Universal Robots URScript: FaiChun_9 Jan_1_arc_1.script

def Machining2():
  # Default parameters:
  global speed_ms = 0.05
  global speed_rads = 0.75
  global accel_mss = 3
  global accel_radss = 1.2
  global blend_radius_m = 0.0003

  # Add subprograms here
  # Start of main program
  # Program generated by RoboDK v5.6.8 for UR10e on 13/01/2025 16:29:17
  # Using nominal kinematics.
  blend_radius_m = 0.0003
  speed_ms = 0.05
  # set_reference(p[0.325000, -0.070000, 0.000000, 0.000000, 0.000000, 0.000000])
  set_tcp(p[0.000000, 0.000000, 0.252000, 0.000000, 0.000000, 0.000000])
  # Show Tool
  movej([0.739676, -0.896584, -2.557623, -1.258182, 1.570796, 2.310473],accel_radss,speed_rads,0,blend_radius_m)
  movel([0.739676, -1.045549, -2.705771, -0.961069, 1.570796, 2.310473],accel_mss,speed_ms,0,blend_radius_m)
  #SetTool1
  #M_RunCode6
  #SetRPM60000
  speed_ms = 0.05
  #M_RunCode3
  movel([0.739676, -1.073443, -2.722043, -0.916902, 1.570796, 2.310473],accel_mss,speed_ms,0,blend_radius_m)
  speed_ms = 0.003
  movel([0.739676, -1.080869, -2.726059, -0.905462, 1.570796, 2.310473],accel_mss,speed_ms,0,blend_radius_m)
  speed_ms = 0.007
  movel([0.521026, -1.435757, -2.529573, -0.747059, 1.570796, 2.091823],accel_mss,speed_ms,0,blend_radius_m)
  movel([0.234867, -1.438478, -2.527424, -0.746487, 1.570796, 1.805663],accel_mss,speed_ms,0,blend_radius_m)
  movel([0.339201, -1.087620, -2.723617, -0.901152, 1.570796, 1.909998],accel_mss,speed_ms,0,blend_radius_m)
  movel([0.739676, -1.080869, -2.726059, -0.905462, 1.570796, 2.310473],accel_mss,speed_ms,0,blend_radius_m)
  speed_ms = 0.003
  movel([0.739676, -1.073443, -2.722043, -0.916902, 1.570796, 2.310473],accel_mss,speed_ms,0,blend_radius_m)
  speed_ms = 0.05
  movel([0.739676, -1.045549, -2.705771, -0.961069, 1.570796, 2.310473],accel_mss,speed_ms,0,blend_radius_m)
  #M_RunCode9
  movel([0.722285, -1.051564, -2.703686, -0.957139, 1.570796, 2.293082],accel_mss,speed_ms,0,blend_radius_m)
  #M_RunCode3
  movel([0.722285, -1.079477, -2.719883, -0.913030, 1.570796, 2.293082],accel_mss,speed_ms,0,blend_radius_m)
  speed_ms = 0.003
  movel([0.722285, -1.086903, -2.723879, -0.901608, 1.570796, 2.293082],accel_mss,speed_ms,0,blend_radius_m)
  speed_ms = 0.007
  movel([0.717716, -1.094057, -2.721252, -0.897081, 1.570796, 2.288512],accel_mss,speed_ms,0,blend_radius_m)
  movel([0.716212, -1.105701, -2.716877, -0.889811, 1.570796, 2.287008],accel_mss,speed_ms,0,blend_radius_m)
  movel([0.711055, -1.104499, -2.717334, -0.890556, 1.570796, 2.281852],accel_mss,speed_ms,0,blend_radius_m)
  movel([0.713896, -1.109311, -2.715495, -0.887583, 1.570796, 2.284692],accel_mss,speed_ms,0,blend_radius_m)
  movel([0.708427, -1.117848, -2.712180, -0.882361, 1.570796, 2.279223],accel_mss,speed_ms,0,blend_radius_m)
  movel([0.707812, -1.118809, -2.711802, -0.881778, 1.570796, 2.278608],accel_mss,speed_ms,0,blend_radius_m)
  movel([0.707378, -1.119487, -2.711535, -0.881367, 1.570796, 2.278174],accel_mss,speed_ms,0,blend_radius_m)
  movel([0.699793, -1.117779, -2.712207, -0.882403, 1.570796, 2.270589],accel_mss,speed_ms,0,blend_radius_m)
  movel([0.704152, -1.110893, -2.714886, -0.886610, 1.570796, 2.274948],accel_mss,speed_ms,0,blend_radius_m)
  movel([0.701466, -1.110302, -2.715114, -0.886973, 1.570796, 2.272262],accel_mss,speed_ms,0,blend_radius_m)
  movel([0.694884, -1.120745, -2.711039, -0.880605, 1.570796, 2.265680],accel_mss,speed_ms,0,blend_radius_m)
  movel([0.705120, -1.123018, -2.710138, -0.879233, 1.570796, 2.275917],accel_mss,speed_ms,0,blend_radius_m)
  movel([0.604989, -1.283325, -2.632898, -0.796166, 1.570796, 2.175785],accel_mss,speed_ms,0,blend_radius_m)
  movel([0.530205, -1.410064, -2.549311, -0.753014, 1.570796, 2.101001],accel_mss,speed_ms,0,blend_radius_m)
  movel([0.521929, -1.408991, -2.550114, -0.753284, 1.570796, 2.092726],accel_mss,speed_ms,0,blend_radius_m)
  movel([0.518334, -1.415415, -2.545281, -0.751692, 1.570796, 2.089130],accel_mss,speed_ms,0,blend_radius_m)
  movel([0.520473, -1.415684, -2.545078, -0.751627, 1.570796, 2.091269],accel_mss,speed_ms,0,blend_radius_m)
  movel([0.522841, -1.411466, -2.548259, -0.752664, 1.570796, 2.093637],accel_mss,speed_ms,0,blend_radius_m)
  movel([0.528942, -1.412267, -2.547657, -0.752465, 1.570796, 2.099738],accel_mss,speed_ms,0,blend_radius_m)
  movel([0.528547, -1.412961, -2.547135, -0.752293, 1.570796, 2.099343],accel_mss,speed_ms,0,blend_radius_m)
  movel([0.528364, -1.413282, -2.546893, -0.752214, 1.570796, 2.099160],accel_mss,speed_ms,0,blend_radius_m)
  movel([0.521314, -1.417954, -2.543354, -0.751080, 1.570796, 2.092111],accel_mss,speed_ms,0,blend_radius_m)
  movec([0.521009, -1.418498, -2.542941, -0.750950, 1.570796, 2.091805],[0.520704, -1.419040, -2.542527, -0.750821, 1.570796, 2.091500],accel_mss,speed_ms,blend_radius_m)
  movec([0.520399, -1.419584, -2.542113, -0.750692, 1.570796, 2.091195],[0.520094, -1.420127, -2.541698, -0.750564, 1.570796, 2.090890],accel_mss,speed_ms,blend_radius_m)
  movel([0.524182, -1.420660, -2.541290, -0.750438, 1.570796, 2.094978],accel_mss,speed_ms,0,blend_radius_m)
  movel([0.520710, -1.426805, -2.536563, -0.749022, 1.570796, 2.091507],accel_mss,speed_ms,0,blend_radius_m)
  movel([0.516647, -1.426280, -2.536969, -0.749140, 1.570796, 2.087443],accel_mss,speed_ms,0,blend_radius_m)
  movel([0.514345, -1.430404, -2.533767, -0.748218, 1.570796, 2.085141],accel_mss,speed_ms,0,blend_radius_m)
  movel([0.508328, -1.429667, -2.534341, -0.748381, 1.570796, 2.079124],accel_mss,speed_ms,0,blend_radius_m)
  movel([0.510606, -1.425534, -2.537545, -0.749310, 1.570796, 2.081402],accel_mss,speed_ms,0,blend_radius_m)
  movel([0.506209, -1.429417, -2.534536, -0.748437, 1.570796, 2.077005],accel_mss,speed_ms,0,blend_radius_m)
  movel([0.501142, -1.428840, -2.534984, -0.748565, 1.570796, 2.071939],accel_mss,speed_ms,0,blend_radius_m)
  movel([0.500651, -1.428783, -2.535029, -0.748578, 1.570796, 2.071447],accel_mss,speed_ms,0,blend_radius_m)
  movel([0.500157, -1.428731, -2.535069, -0.748589, 1.570796, 2.070953],accel_mss,speed_ms,0,blend_radius_m)
  movel([0.503495, -1.422587, -2.539814, -0.749988, 1.570796, 2.074291],accel_mss,speed_ms,0,blend_radius_m)
  movel([0.507609, -1.423054, -2.539455, -0.749880, 1.570796, 2.078405],accel_mss,speed_ms,0,blend_radius_m)
  movel([0.508797, -1.420891, -2.541114, -0.750384, 1.570796, 2.079593],accel_mss,speed_ms,0,blend_radius_m)
  movel([0.502532, -1.420185, -2.541654, -0.750550, 1.570796, 2.073328],accel_mss,speed_ms,0,blend_radius_m)
  movel([0.498030, -1.428499, -2.535249, -0.748641, 1.570796, 2.068827],accel_mss,speed_ms,0,blend_radius_m)
  movel([0.497523, -1.428447, -2.535290, -0.748653, 1.570796, 2.068319],accel_mss,speed_ms,0,blend_radius_m)
  movel([0.497042, -1.428395, -2.535329, -0.748664, 1.570796, 2.067838],accel_mss,speed_ms,0,blend_radius_m)
  movel([0.383251, -1.423074, -2.539440, -0.749875, 1.570796, 1.954047],accel_mss,speed_ms,0,blend_radius_m)
  movel([0.263080, -1.430856, -2.533414, -0.748118, 1.570796, 1.833877],accel_mss,speed_ms,0,blend_radius_m)
  movel([0.265517, -1.422588, -2.539813, -0.749988, 1.570796, 1.836314],accel_mss,speed_ms,0,blend_radius_m)
  movel([0.258622, -1.423422, -2.539172, -0.749794, 1.570796, 1.829418],accel_mss,speed_ms,0,blend_radius_m)
  movel([0.257999, -1.425574, -2.537514, -0.749301, 1.570796, 1.828796],accel_mss,speed_ms,0,blend_radius_m)
  movel([0.262529, -1.425022, -2.537940, -0.749427, 1.570796, 1.833326],accel_mss,speed_ms,0,blend_radius_m)
  movel([0.260738, -1.431127, -2.533203, -0.748059, 1.570796, 1.831534],accel_mss,speed_ms,0,blend_radius_m)
  movel([0.259655, -1.431256, -2.533102, -0.748031, 1.570796, 1.830452],accel_mss,speed_ms,0,blend_radius_m)
  movel([0.255252, -1.427829, -2.535769, -0.748791, 1.570796, 1.826048],accel_mss,speed_ms,0,blend_radius_m)
  movel([0.252906, -1.428125, -2.535539, -0.748725, 1.570796, 1.823702],accel_mss,speed_ms,0,blend_radius_m)
  movel([0.251743, -1.432228, -2.532342, -0.747818, 1.570796, 1.822539],accel_mss,speed_ms,0,blend_radius_m)
  movel([0.245076, -1.433089, -2.531668, -0.747631, 1.570796, 1.815873],accel_mss,speed_ms,0,blend_radius_m)
  movel([0.246206, -1.428996, -2.534863, -0.748530, 1.570796, 1.817002],accel_mss,speed_ms,0,blend_radius_m)
  movel([0.243345, -1.423504, -2.539109, -0.749776, 1.570796, 1.814141],accel_mss,speed_ms,0,blend_radius_m)
  movel([0.247902, -1.422884, -2.539586, -0.749919, 1.570796, 1.818698],accel_mss,speed_ms,0,blend_radius_m)
  movel([0.248502, -1.420729, -2.541238, -0.750422, 1.570796, 1.819298],accel_mss,speed_ms,0,blend_radius_m)
  movel([0.243934, -1.421351, -2.540762, -0.750276, 1.570796, 1.814730],accel_mss,speed_ms,0,blend_radius_m)
  movel([0.245350, -1.416182, -2.544701, -0.751507, 1.570796, 1.816147],accel_mss,speed_ms,0,blend_radius_m)
  movel([0.252445, -1.414242, -2.546169, -0.751979, 1.570796, 1.823242],accel_mss,speed_ms,0,blend_radius_m)
  movel([0.251262, -1.418432, -2.542991, -0.750966, 1.570796, 1.822058],accel_mss,speed_ms,0,blend_radius_m)
  movel([0.253639, -1.418118, -2.543230, -0.751041, 1.570796, 1.824436],accel_mss,speed_ms,0,blend_radius_m)
  movel([0.255455, -1.411739, -2.548054, -0.752596, 1.570796, 1.826251],accel_mss,speed_ms,0,blend_radius_m)
  movel([0.246231, -1.412992, -2.547111, -0.752286, 1.570796, 1.817027],accel_mss,speed_ms,0,blend_radius_m)
  movel([0.282412, -1.287409, -2.630540, -0.794439, 1.570796, 1.853209],accel_mss,speed_ms,0,blend_radius_m)
  movel([0.331289, -1.130759, -2.707034, -0.874596, 1.570796, 1.902085],accel_mss,speed_ms,0,blend_radius_m)
  movel([0.331811, -1.129158, -2.707681, -0.875550, 1.570796, 1.902607],accel_mss,speed_ms,0,blend_radius_m)
  movel([0.344365, -1.126524, -2.708739, -0.877125, 1.570796, 1.915161],accel_mss,speed_ms,0,blend_radius_m)
  movel([0.347816, -1.116232, -2.712812, -0.883345, 1.570796, 1.918612],accel_mss,speed_ms,0,blend_radius_m)
  movel([0.344526, -1.116917, -2.712545, -0.882928, 1.570796, 1.915323],accel_mss,speed_ms,0,blend_radius_m)
  movel([0.342270, -1.123698, -2.709868, -0.878823, 1.570796, 1.913066],accel_mss,speed_ms,0,blend_radius_m)
  movel([0.332951, -1.125669, -2.709082, -0.877638, 1.570796, 1.903747],accel_mss,speed_ms,0,blend_radius_m)
  movel([0.333474, -1.124054, -2.709726, -0.878609, 1.570796, 1.904271],accel_mss,speed_ms,0,blend_radius_m)
  movel([0.342570, -1.114276, -2.713575, -0.884538, 1.570796, 1.913366],accel_mss,speed_ms,0,blend_radius_m)
  movel([0.343748, -1.110711, -2.714956, -0.886722, 1.570796, 1.914545],accel_mss,speed_ms,0,blend_radius_m)
  movel([0.340718, -1.101853, -2.718336, -0.892200, 1.570796, 1.911515],accel_mss,speed_ms,0,blend_radius_m)
  movel([0.347166, -1.100432, -2.718872, -0.893085, 1.570796, 1.917962],accel_mss,speed_ms,0,blend_radius_m)
  movel([0.349516, -1.093391, -2.721498, -0.897500, 1.570796, 1.920312],accel_mss,speed_ms,0,blend_radius_m)
  movel([0.359125, -1.091319, -2.722262, -0.898808, 1.570796, 1.929921],accel_mss,speed_ms,0,blend_radius_m)
  movel([0.356708, -1.098395, -2.719636, -0.894358, 1.570796, 1.927504],accel_mss,speed_ms,0,blend_radius_m)
  movec([0.357543, -1.098221, -2.719701, -0.894467, 1.570796, 1.928339],[0.358378, -1.098047, -2.719766, -0.894576, 1.570796, 1.929174],accel_mss,speed_ms,blend_radius_m)
  movec([0.359213, -1.097874, -2.719831, -0.894684, 1.570796, 1.930010],[0.360048, -1.097701, -2.719896, -0.894792, 1.570796, 1.930844],accel_mss,speed_ms,blend_radius_m)
  movel([0.362489, -1.090612, -2.722522, -0.899255, 1.570796, 1.933285],accel_mss,speed_ms,0,blend_radius_m)
  movel([0.372081, -1.088653, -2.723240, -0.900496, 1.570796, 1.942877],accel_mss,speed_ms,0,blend_radius_m)
  movel([0.368381, -1.099168, -2.719347, -0.893875, 1.570796, 1.939178],accel_mss,speed_ms,0,blend_radius_m)
  movel([0.361972, -1.100448, -2.718866, -0.893075, 1.570796, 1.932768],accel_mss,speed_ms,0,blend_radius_m)
  movel([0.360716, -1.104083, -2.717492, -0.890814, 1.570796, 1.931512],accel_mss,speed_ms,0,blend_radius_m)
  movel([0.370416, -1.102170, -2.718216, -0.892002, 1.570796, 1.941212],accel_mss,speed_ms,0,blend_radius_m)
  movel([0.375438, -1.087987, -2.723483, -0.900919, 1.570796, 1.946234],accel_mss,speed_ms,0,blend_radius_m)
  movel([0.546051, -1.068879, -2.730296, -0.913214, 1.570796, 2.116847],accel_mss,speed_ms,0,blend_radius_m)
  movel([0.701149, -1.082254, -2.725561, -0.904574, 1.570796, 2.271946],accel_mss,speed_ms,0,blend_radius_m)
  movel([0.692244, -1.096648, -2.720289, -0.895452, 1.570796, 2.263040],accel_mss,speed_ms,0,blend_radius_m)
  movel([0.700259, -1.098274, -2.719681, -0.894433, 1.570796, 2.271055],accel_mss,speed_ms,0,blend_radius_m)
  movel([0.702567, -1.094590, -2.721054, -0.896745, 1.570796, 2.273363],accel_mss,speed_ms,0,blend_radius_m)
  movel([0.697284, -1.093499, -2.721458, -0.897432, 1.570796, 2.268081],accel_mss,speed_ms,0,blend_radius_m)
  movel([0.703923, -1.082833, -2.725353, -0.904204, 1.570796, 2.274720],accel_mss,speed_ms,0,blend_radius_m)
  movel([0.704189, -1.082887, -2.725333, -0.904169, 1.570796, 2.274985],accel_mss,speed_ms,0,blend_radius_m)
  movel([0.705203, -1.083098, -2.725257, -0.904034, 1.570796, 2.275999],accel_mss,speed_ms,0,blend_radius_m)
  movel([0.711781, -1.084505, -2.724749, -0.903135, 1.570796, 2.282578],accel_mss,speed_ms,0,blend_radius_m)
  movel([0.707252, -1.091700, -2.722122, -0.898567, 1.570796, 2.278048],accel_mss,speed_ms,0,blend_radius_m)
  movel([0.709979, -1.092296, -2.721902, -0.898191, 1.570796, 2.280775],accel_mss,speed_ms,0,blend_radius_m)
  movel([0.722285, -1.086903, -2.723879, -0.901608, 1.570796, 2.293082],accel_mss,speed_ms,0,blend_radius_m)
  speed_ms = 0.003
  movel([0.722285, -1.079477, -2.719883, -0.913030, 1.570796, 2.293082],accel_mss,speed_ms,0,blend_radius_m)
  speed_ms = 0.05
  movel([0.722285, -1.051564, -2.703686, -0.957139, 1.570796, 2.293082],accel_mss,speed_ms,0,blend_radius_m)
  #M_RunCode9
  movel([0.397634, -1.094593, -2.687861, -0.929935, 1.570796, 1.968430],accel_mss,speed_ms,0,blend_radius_m)
  #M_RunCode3
  movel([0.397634, -1.122537, -2.703510, -0.886342, 1.570796, 1.968430],accel_mss,speed_ms,0,blend_radius_m)
  speed_ms = 0.003
  movel([0.397634, -1.129941, -2.707365, -0.875083, 1.570796, 1.968430],accel_mss,speed_ms,0,blend_radius_m)
  speed_ms = 0.007
  movec([0.397337, -1.130959, -2.706953, -0.874477, 1.570796, 1.968133],[0.396949, -1.131993, -2.706534, -0.873862, 1.570796, 1.967745],accel_mss,speed_ms,blend_radius_m)
  movec([0.396255, -1.133449, -2.705942, -0.872998, 1.570796, 1.967051],[0.395394, -1.134891, -2.705353, -0.872144, 1.570796, 1.966190],accel_mss,speed_ms,blend_radius_m)
  movec([0.394595, -1.136025, -2.704889, -0.871475, 1.570796, 1.965391],[0.393717, -1.137121, -2.704440, -0.870829, 1.570796, 1.964513],accel_mss,speed_ms,blend_radius_m)
  movec([0.392871, -1.138072, -2.704048, -0.870269, 1.570796, 1.963667],[0.391984, -1.138986, -2.703672, -0.869732, 1.570796, 1.962780],accel_mss,speed_ms,blend_radius_m)
  movec([0.390895, -1.140016, -2.703246, -0.869127, 1.570796, 1.961691],[0.389771, -1.140994, -2.702841, -0.868555, 1.570796, 1.960567],accel_mss,speed_ms,blend_radius_m)
  movec([0.388667, -1.141870, -2.702477, -0.868042, 1.570796, 1.959464],[0.387540, -1.142678, -2.702141, -0.867570, 1.570796, 1.958336],accel_mss,speed_ms,blend_radius_m)
  movec([0.386309, -1.143464, -2.701813, -0.867112, 1.570796, 1.957105],[0.385068, -1.144158, -2.701523, -0.866707, 1.570796, 1.955864],accel_mss,speed_ms,blend_radius_m)
  movel([0.384283, -1.144545, -2.701362, -0.866482, 1.570796, 1.955080],accel_mss,speed_ms,0,blend_radius_m)
  movec([0.382774, -1.145210, -2.701083, -0.866096, 1.570796, 1.953570],[0.381275, -1.145785, -2.700842, -0.865762, 1.570796, 1.952072],accel_mss,speed_ms,blend_radius_m)
  movec([0.379746, -1.146284, -2.700633, -0.865472, 1.570796, 1.950543],[0.378243, -1.146680, -2.700466, -0.865242, 1.570796, 1.949039],accel_mss,speed_ms,blend_radius_m)
  movel([0.377080, -1.146932, -2.700360, -0.865097, 1.570796, 1.947876],accel_mss,speed_ms,0,blend_radius_m)
  movec([0.375723, -1.147196, -2.700249, -0.864943, 1.570796, 1.946520],[0.374377, -1.147434, -2.700149, -0.864806, 1.570796, 1.945173],accel_mss,speed_ms,blend_radius_m)
  movec([0.372777, -1.147687, -2.700043, -0.864660, 1.570796, 1.943574],[0.371187, -1.147915, -2.699946, -0.864527, 1.570796, 1.941984],accel_mss,speed_ms,blend_radius_m)
  movec([0.368942, -1.148277, -2.699794, -0.864318, 1.570796, 1.939738],[0.366679, -1.148691, -2.699619, -0.864079, 1.570796, 1.937475],accel_mss,speed_ms,blend_radius_m)
  movec([0.365810, -1.148867, -2.699545, -0.863977, 1.570796, 1.936606],[0.364936, -1.149059, -2.699464, -0.863867, 1.570796, 1.935733],accel_mss,speed_ms,blend_radius_m)
  movel([0.364507, -1.149159, -2.699421, -0.863809, 1.570796, 1.935303],accel_mss,speed_ms,0,blend_radius_m)
  movec([0.363623, -1.149389, -2.699324, -0.863676, 1.570796, 1.934419],[0.362729, -1.149654, -2.699212, -0.863523, 1.570796, 1.933525],accel_mss,speed_ms,blend_radius_m)
  movec([0.361556, -1.150059, -2.699040, -0.863290, 1.570796, 1.932352],[0.360373, -1.150529, -2.698841, -0.863019, 1.570796, 1.931169],accel_mss,speed_ms,blend_radius_m)
  movel([0.359060, -1.151121, -2.698590, -0.862678, 1.570796, 1.929857],accel_mss,speed_ms,0,blend_radius_m)
  movel([0.357816, -1.151769, -2.698314, -0.862306, 1.570796, 1.928612],accel_mss,speed_ms,0,blend_radius_m)
  movec([0.356426, -1.152631, -2.697947, -0.861811, 1.570796, 1.927223],[0.355071, -1.153621, -2.697525, -0.861244, 1.570796, 1.925867],accel_mss,speed_ms,blend_radius_m)
  movec([0.354412, -1.154159, -2.697294, -0.860936, 1.570796, 1.925208],[0.353768, -1.154723, -2.697053, -0.860613, 1.570796, 1.924564],accel_mss,speed_ms,blend_radius_m)
  movel([0.353988, -1.155027, -2.696922, -0.860439, 1.570796, 1.924784],accel_mss,speed_ms,0,blend_radius_m)
  movel([0.354205, -1.155333, -2.696791, -0.860265, 1.570796, 1.925001],accel_mss,speed_ms,0,blend_radius_m)
  movel([0.354363, -1.155556, -2.696696, -0.860137, 1.570796, 1.925159],accel_mss,speed_ms,0,blend_radius_m)
  movec([0.355113, -1.156538, -2.696274, -0.859578, 1.570796, 1.925909],[0.355924, -1.157459, -2.695877, -0.859053, 1.570796, 1.926721],accel_mss,speed_ms,blend_radius_m)
  movec([0.356629, -1.158142, -2.695582, -0.858665, 1.570796, 1.927425],[0.357388, -1.158766, -2.695312, -0.858310, 1.570796, 1.928184],accel_mss,speed_ms,blend_radius_m)
  movec([0.358002, -1.159195, -2.695127, -0.858067, 1.570796, 1.928799],[0.358655, -1.159578, -2.694961, -0.857850, 1.570796, 1.929451],accel_mss,speed_ms,blend_radius_m)
  movec([0.359290, -1.159888, -2.694826, -0.857674, 1.570796, 1.930086],[0.359960, -1.160152, -2.694712, -0.857525, 1.570796, 1.930756],accel_mss,speed_ms,blend_radius_m)
  movec([0.360746, -1.160381, -2.694612, -0.857396, 1.570796, 1.931543],[0.361580, -1.160537, -2.694545, -0.857308, 1.570796, 1.932376],accel_mss,speed_ms,blend_radius_m)
  movel([0.362491, -1.160615, -2.694511, -0.857263, 1.570796, 1.933287],accel_mss,speed_ms,0,blend_radius_m)
  movec([0.363505, -1.160603, -2.694516, -0.857270, 1.570796, 1.934301],[0.364559, -1.160501, -2.694560, -0.857328, 1.570796, 1.935355],accel_mss,speed_ms,blend_radius_m)
  movec([0.365638, -1.160307, -2.694644, -0.857437, 1.570796, 1.936435],[0.366749, -1.160013, -2.694772, -0.857604, 1.570796, 1.937545],accel_mss,speed_ms,blend_radius_m)
  movec([0.368362, -1.159420, -2.695029, -0.857940, 1.570796, 1.939159],[0.369995, -1.158626, -2.695373, -0.858390, 1.570796, 1.940791],accel_mss,speed_ms,blend_radius_m)
  movec([0.371113, -1.157977, -2.695653, -0.858759, 1.570796, 1.941909],[0.372219, -1.157253, -2.695966, -0.859170, 1.570796, 1.943015],accel_mss,speed_ms,blend_radius_m)
  movel([0.360789, -1.167387, -2.691545, -0.853457, 1.570796, 1.931585],accel_mss,speed_ms,0,blend_radius_m)
  movel([0.344914, -1.145108, -2.701126, -0.866155, 1.570796, 1.915710],accel_mss,speed_ms,0,blend_radius_m)
  movel([0.346071, -1.144040, -2.701573, -0.866776, 1.570796, 1.916867],accel_mss,speed_ms,0,blend_radius_m)
  movec([0.347403, -1.142893, -2.702051, -0.867445, 1.570796, 1.918199],[0.348790, -1.141858, -2.702482, -0.868049, 1.570796, 1.919586],accel_mss,speed_ms,blend_radius_m)
  movec([0.349938, -1.141112, -2.702792, -0.868485, 1.570796, 1.920734],[0.351098, -1.140448, -2.703067, -0.868874, 1.570796, 1.921894],accel_mss,speed_ms,blend_radius_m)
  movec([0.351876, -1.140050, -2.703232, -0.869107, 1.570796, 1.922673],[0.352654, -1.139687, -2.703382, -0.869320, 1.570796, 1.923450],accel_mss,speed_ms,blend_radius_m)
  movec([0.354924, -1.138754, -2.703767, -0.869868, 1.570796, 1.925721],[0.357169, -1.137991, -2.704082, -0.870316, 1.570796, 1.927965],accel_mss,speed_ms,blend_radius_m)
  movec([0.358472, -1.137621, -2.704234, -0.870534, 1.570796, 1.929269],[0.359759, -1.137311, -2.704362, -0.870717, 1.570796, 1.930556],accel_mss,speed_ms,blend_radius_m)
  movec([0.360451, -1.137162, -2.704423, -0.870805, 1.570796, 1.931247],[0.361141, -1.137017, -2.704482, -0.870890, 1.570796, 1.931938],accel_mss,speed_ms,blend_radius_m)
  movec([0.362865, -1.136681, -2.704620, -0.871088, 1.570796, 1.933661],[0.364580, -1.136371, -2.704747, -0.871271, 1.570796, 1.935376],accel_mss,speed_ms,blend_radius_m)
  movec([0.366768, -1.136001, -2.704899, -0.871489, 1.570796, 1.937564],[0.368948, -1.135654, -2.705041, -0.871694, 1.570796, 1.939744],accel_mss,speed_ms,blend_radius_m)
  movec([0.371841, -1.135226, -2.705217, -0.871947, 1.570796, 1.942637],[0.374749, -1.134761, -2.705407, -0.872222, 1.570796, 1.945545],accel_mss,speed_ms,blend_radius_m)
  movec([0.375820, -1.134576, -2.705482, -0.872331, 1.570796, 1.946616],[0.376896, -1.134377, -2.705563, -0.872449, 1.570796, 1.947692],accel_mss,speed_ms,blend_radius_m)
  movel([0.377425, -1.134273, -2.705606, -0.872510, 1.570796, 1.948222],accel_mss,speed_ms,0,blend_radius_m)
  movec([0.379248, -1.133855, -2.705776, -0.872758, 1.570796, 1.950044],[0.381104, -1.133317, -2.705996, -0.873076, 1.570796, 1.951900],accel_mss,speed_ms,blend_radius_m)
  movec([0.382534, -1.132825, -2.706196, -0.873368, 1.570796, 1.953331],[0.383978, -1.132256, -2.706427, -0.873706, 1.570796, 1.954775],accel_mss,speed_ms,blend_radius_m)
  movec([0.385185, -1.131706, -2.706650, -0.874032, 1.570796, 1.955982],[0.386396, -1.131064, -2.706911, -0.874414, 1.570796, 1.957192],accel_mss,speed_ms,blend_radius_m)
  movec([0.387452, -1.130417, -2.707172, -0.874799, 1.570796, 1.958248],[0.388493, -1.129686, -2.707468, -0.875235, 1.570796, 1.959289],accel_mss,speed_ms,blend_radius_m)
  movec([0.389177, -1.129152, -2.707683, -0.875554, 1.570796, 1.959973],[0.389847, -1.128585, -2.707912, -0.875892, 1.570796, 1.960643],accel_mss,speed_ms,blend_radius_m)
  movec([0.390510, -1.127977, -2.708156, -0.876256, 1.570796, 1.961306],[0.391154, -1.127344, -2.708410, -0.876634, 1.570796, 1.961951],accel_mss,speed_ms,blend_radius_m)
  movel([0.392177, -1.126228, -2.708858, -0.877303, 1.570796, 1.962973],accel_mss,speed_ms,0,blend_radius_m)
  movel([0.393116, -1.125005, -2.709347, -0.878037, 1.570796, 1.963912],accel_mss,speed_ms,0,blend_radius_m)
  movel([0.393830, -1.123845, -2.709809, -0.878734, 1.570796, 1.964626],accel_mss,speed_ms,0,blend_radius_m)
  movel([0.394302, -1.122851, -2.710205, -0.879333, 1.570796, 1.965098],accel_mss,speed_ms,0,blend_radius_m)
  movel([0.394449, -1.122460, -2.710360, -0.879569, 1.570796, 1.965245],accel_mss,speed_ms,0,blend_radius_m)
  movec([0.394689, -1.121685, -2.710667, -0.880037, 1.570796, 1.965485],[0.394858, -1.120928, -2.710966, -0.880494, 1.570796, 1.965654],accel_mss,speed_ms,blend_radius_m)
  movec([0.394959, -1.119764, -2.711426, -0.881199, 1.570796, 1.965755],[0.394824, -1.118725, -2.711835, -0.881829, 1.570796, 1.965621],accel_mss,speed_ms,blend_radius_m)
  movel([0.394458, -1.117809, -2.712195, -0.882385, 1.570796, 1.965254],accel_mss,speed_ms,0,blend_radius_m)
  movec([0.394177, -1.117385, -2.712361, -0.882643, 1.570796, 1.964973],[0.393846, -1.117007, -2.712509, -0.882872, 1.570796, 1.964643],accel_mss,speed_ms,blend_radius_m)
  movel([0.393215, -1.116570, -2.712680, -0.883139, 1.570796, 1.964012],accel_mss,speed_ms,0,blend_radius_m)
  movel([0.392747, -1.116425, -2.712737, -0.883227, 1.570796, 1.963544],accel_mss,speed_ms,0,blend_radius_m)
  movel([0.392465, -1.116395, -2.712749, -0.883245, 1.570796, 1.963261],accel_mss,speed_ms,0,blend_radius_m)
  movel([0.391761, -1.116466, -2.712721, -0.883202, 1.570796, 1.962558],accel_mss,speed_ms,0,blend_radius_m)
  movel([0.391189, -1.116670, -2.712641, -0.883078, 1.570796, 1.961986],accel_mss,speed_ms,0,blend_radius_m)
  movel([0.390941, -1.116802, -2.712590, -0.882998, 1.570796, 1.961738],accel_mss,speed_ms,0,blend_radius_m)
  movel([0.390599, -1.117028, -2.712501, -0.882860, 1.570796, 1.961395],accel_mss,speed_ms,0,blend_radius_m)
  movel([0.390249, -1.117314, -2.712389, -0.882686, 1.570796, 1.961045],accel_mss,speed_ms,0,blend_radius_m)
  movel([0.390069, -1.117494, -2.712318, -0.882576, 1.570796, 1.960865],accel_mss,speed_ms,0,blend_radius_m)
  movel([0.389660, -1.118019, -2.712112, -0.882257, 1.570796, 1.960456],accel_mss,speed_ms,0,blend_radius_m)
  movel([0.389214, -1.118739, -2.711829, -0.881820, 1.570796, 1.960010],accel_mss,speed_ms,0,blend_radius_m)
  movel([0.389063, -1.119009, -2.711723, -0.881657, 1.570796, 1.959860],accel_mss,speed_ms,0,blend_radius_m)
  movel([0.388430, -1.120085, -2.711299, -0.881004, 1.570796, 1.959226],accel_mss,speed_ms,0,blend_radius_m)
  movel([0.388001, -1.120712, -2.711052, -0.880625, 1.570796, 1.958798],accel_mss,speed_ms,0,blend_radius_m)
  movel([0.387698, -1.121101, -2.710898, -0.880390, 1.570796, 1.958494],accel_mss,speed_ms,0,blend_radius_m)
  movel([0.386944, -1.121913, -2.710577, -0.879899, 1.570796, 1.957740],accel_mss,speed_ms,0,blend_radius_m)
  movel([0.385868, -1.122888, -2.710190, -0.879311, 1.570796, 1.956664],accel_mss,speed_ms,0,blend_radius_m)
  movel([0.384591, -1.123812, -2.709823, -0.878755, 1.570796, 1.955387],accel_mss,speed_ms,0,blend_radius_m)
  movel([0.383635, -1.124316, -2.709622, -0.878451, 1.570796, 1.954431],accel_mss,speed_ms,0,blend_radius_m)
  movel([0.382614, -1.124643, -2.709491, -0.878255, 1.570796, 1.953411],accel_mss,speed_ms,0,blend_radius_m)
  movel([0.381863, -1.124736, -2.709454, -0.878199, 1.570796, 1.952660],accel_mss,speed_ms,0,blend_radius_m)
  movel([0.381227, -1.124716, -2.709462, -0.878211, 1.570796, 1.952024],accel_mss,speed_ms,0,blend_radius_m)
  movec([0.380479, -1.124561, -2.709524, -0.878304, 1.570796, 1.951276],[0.379833, -1.124259, -2.709645, -0.878486, 1.570796, 1.950629],accel_mss,speed_ms,blend_radius_m)
  movec([0.379397, -1.123934, -2.709774, -0.878681, 1.570796, 1.950193],[0.379025, -1.123539, -2.709931, -0.878919, 1.570796, 1.949822],accel_mss,speed_ms,blend_radius_m)
  movel([0.378826, -1.123266, -2.710040, -0.879083, 1.570796, 1.949623],accel_mss,speed_ms,0,blend_radius_m)
  movec([0.378562, -1.122785, -2.710231, -0.879373, 1.570796, 1.949358],[0.378361, -1.122252, -2.710442, -0.879695, 1.570796, 1.949157],accel_mss,speed_ms,blend_radius_m)
  movec([0.378238, -1.121691, -2.710665, -0.880033, 1.570796, 1.949035],[0.378194, -1.121081, -2.710906, -0.880402, 1.570796, 1.948990],accel_mss,speed_ms,blend_radius_m)
  movel([0.378257, -1.120171, -2.711265, -0.880952, 1.570796, 1.949053],accel_mss,speed_ms,0,blend_radius_m)
  movel([0.378471, -1.119188, -2.711653, -0.881548, 1.570796, 1.949268],accel_mss,speed_ms,0,blend_radius_m)
  movel([0.378817, -1.118259, -2.712018, -0.882112, 1.570796, 1.949614],accel_mss,speed_ms,0,blend_radius_m)
  movec([0.379196, -1.117536, -2.712302, -0.882551, 1.570796, 1.949992],[0.379662, -1.116824, -2.712581, -0.882984, 1.570796, 1.950459],accel_mss,speed_ms,blend_radius_m)
  movel([0.380536, -1.115764, -2.712995, -0.883630, 1.570796, 1.951332],accel_mss,speed_ms,0,blend_radius_m)
  movel([0.381267, -1.115031, -2.713281, -0.884077, 1.570796, 1.952063],accel_mss,speed_ms,0,blend_radius_m)
  movel([0.381574, -1.114752, -2.713390, -0.884247, 1.570796, 1.952371],accel_mss,speed_ms,0,blend_radius_m)
  movec([0.382261, -1.114173, -2.713615, -0.884601, 1.570796, 1.953057],[0.382967, -1.113639, -2.713823, -0.884927, 1.570796, 1.953763],accel_mss,speed_ms,blend_radius_m)
  movel([0.384108, -1.112917, -2.714103, -0.885369, 1.570796, 1.954904],accel_mss,speed_ms,0,blend_radius_m)
  movec([0.384953, -1.112494, -2.714267, -0.885628, 1.570796, 1.955750],[0.385789, -1.112171, -2.714392, -0.885826, 1.570796, 1.956585],accel_mss,speed_ms,blend_radius_m)
  movec([0.386666, -1.111937, -2.714483, -0.885970, 1.570796, 1.957462],[0.387505, -1.111814, -2.714530, -0.886045, 1.570796, 1.958301],accel_mss,speed_ms,blend_radius_m)
  movec([0.388225, -1.111790, -2.714539, -0.886060, 1.570796, 1.959022],[0.388911, -1.111835, -2.714522, -0.886032, 1.570796, 1.959707],accel_mss,speed_ms,blend_radius_m)
  movel([0.389300, -1.111895, -2.714499, -0.885995, 1.570796, 1.960097],accel_mss,speed_ms,0,blend_radius_m)
  movec([0.390012, -1.112053, -2.714438, -0.885899, 1.570796, 1.960808],[0.390685, -1.112268, -2.714354, -0.885766, 1.570796, 1.961481],accel_mss,speed_ms,blend_radius_m)
  movec([0.391772, -1.112759, -2.714164, -0.885465, 1.570796, 1.962568],[0.392753, -1.113384, -2.713922, -0.885083, 1.570796, 1.963549],accel_mss,speed_ms,blend_radius_m)
  movec([0.393548, -1.114044, -2.713665, -0.884680, 1.570796, 1.964345],[0.394269, -1.114783, -2.713378, -0.884228, 1.570796, 1.965065],accel_mss,speed_ms,blend_radius_m)
  movec([0.394949, -1.115628, -2.713048, -0.883712, 1.570796, 1.965746],[0.395564, -1.116535, -2.712694, -0.883160, 1.570796, 1.966360],accel_mss,speed_ms,blend_radius_m)
  movec([0.396177, -1.117613, -2.712272, -0.882505, 1.570796, 1.966973],[0.396716, -1.118751, -2.711825, -0.881813, 1.570796, 1.967512],accel_mss,speed_ms,blend_radius_m)
  movec([0.397337, -1.120472, -2.711147, -0.880770, 1.570796, 1.968133],[0.397782, -1.122317, -2.710416, -0.879655, 1.570796, 1.968578],accel_mss,speed_ms,blend_radius_m)
  movec([0.398010, -1.124002, -2.709747, -0.878640, 1.570796, 1.968807],[0.398085, -1.125773, -2.709040, -0.877576, 1.570796, 1.968881],accel_mss,speed_ms,blend_radius_m)
  movec([0.398059, -1.126856, -2.708607, -0.876927, 1.570796, 1.968855],[0.397980, -1.127962, -2.708162, -0.876264, 1.570796, 1.968776],accel_mss,speed_ms,blend_radius_m)
  movec([0.397847, -1.128938, -2.707770, -0.875682, 1.570796, 1.968644],[0.397634, -1.129941, -2.707365, -0.875083, 1.570796, 1.968430],accel_mss,speed_ms,blend_radius_m)
  speed_ms = 0.003
  movel([0.397634, -1.122537, -2.703510, -0.886342, 1.570796, 1.968430],accel_mss,speed_ms,0,blend_radius_m)
  speed_ms = 0.05
  movel([0.397634, -1.094593, -2.687861, -0.929935, 1.570796, 1.968430],accel_mss,speed_ms,0,blend_radius_m)
  #M_RunCode9
  movel([0.402885, -1.112693, -2.680709, -0.918987, 1.570796, 1.973681],accel_mss,speed_ms,0,blend_radius_m)
  #M_RunCode3
  movel([0.402885, -1.140599, -2.696125, -0.875666, 1.570796, 1.973681],accel_mss,speed_ms,0,blend_radius_m)
  speed_ms = 0.003
  movel([0.402885, -1.147981, -2.699919, -0.864490, 1.570796, 1.973681],accel_mss,speed_ms,0,blend_radius_m)
  speed_ms = 0.007
  movec([0.403566, -1.147510, -2.700117, -0.864762, 1.570796, 1.974362],[0.404251, -1.147054, -2.700309, -0.865026, 1.570796, 1.975047],accel_mss,speed_ms,blend_radius_m)
  movel([0.404789, -1.146708, -2.700454, -0.865226, 1.570796, 1.975586],accel_mss,speed_ms,0,blend_radius_m)
  movec([0.405462, -1.146300, -2.700626, -0.865463, 1.570796, 1.976258],[0.406137, -1.145917, -2.700787, -0.865685, 1.570796, 1.976933],accel_mss,speed_ms,blend_radius_m)
  movec([0.406888, -1.145535, -2.700947, -0.865907, 1.570796, 1.977685],[0.407637, -1.145211, -2.701083, -0.866095, 1.570796, 1.978433],accel_mss,speed_ms,blend_radius_m)
  movel([0.408830, -1.144850, -2.701234, -0.866305, 1.570796, 1.979626],accel_mss,speed_ms,0,blend_radius_m)
  movel([0.409773, -1.144785, -2.701261, -0.866343, 1.570796, 1.980569],accel_mss,speed_ms,0,blend_radius_m)
  movec([0.410338, -1.144915, -2.701207, -0.866267, 1.570796, 1.981135],[0.410790, -1.145199, -2.701088, -0.866102, 1.570796, 1.981586],accel_mss,speed_ms,blend_radius_m)
  movec([0.411125, -1.145616, -2.700913, -0.865860, 1.570796, 1.981921],[0.411335, -1.146140, -2.700693, -0.865556, 1.570796, 1.982132],accel_mss,speed_ms,blend_radius_m)
  movel([0.411361, -1.147181, -2.700256, -0.864952, 1.570796, 1.982157],accel_mss,speed_ms,0,blend_radius_m)
  movel([0.411126, -1.148050, -2.699889, -0.864449, 1.570796, 1.981923],accel_mss,speed_ms,0,blend_radius_m)
  movel([0.410592, -1.149189, -2.699409, -0.863792, 1.570796, 1.981389],accel_mss,speed_ms,0,blend_radius_m)
  movel([0.410020, -1.150105, -2.699021, -0.863263, 1.570796, 1.980816],accel_mss,speed_ms,0,blend_radius_m)
  movel([0.409109, -1.151337, -2.698498, -0.862554, 1.570796, 1.979905],accel_mss,speed_ms,0,blend_radius_m)
  movec([0.408427, -1.152157, -2.698149, -0.862083, 1.570796, 1.979223],[0.407718, -1.152958, -2.697808, -0.861624, 1.570796, 1.978514],accel_mss,speed_ms,blend_radius_m)
  movel([0.406839, -1.153895, -2.697407, -0.861087, 1.570796, 1.977636],accel_mss,speed_ms,0,blend_radius_m)
  movec([0.405648, -1.155117, -2.696884, -0.860388, 1.570796, 1.976444],[0.404438, -1.156317, -2.696369, -0.859703, 1.570796, 1.975234],accel_mss,speed_ms,blend_radius_m)
  movec([0.402822, -1.157867, -2.695701, -0.858821, 1.570796, 1.973618],[0.401189, -1.159388, -2.695043, -0.857958, 1.570796, 1.971985],accel_mss,speed_ms,blend_radius_m)
  movec([0.398900, -1.161468, -2.694140, -0.856781, 1.570796, 1.969696],[0.396598, -1.163513, -2.693247, -0.855629, 1.570796, 1.967394],accel_mss,speed_ms,blend_radius_m)
  movec([0.393071, -1.166572, -2.691904, -0.853912, 1.570796, 1.963867],[0.389532, -1.169574, -2.690577, -0.852238, 1.570796, 1.960328],accel_mss,speed_ms,blend_radius_m)
  movec([0.387356, -1.171381, -2.689773, -0.851234, 1.570796, 1.958153],[0.385172, -1.173159, -2.688980, -0.850250, 1.570796, 1.955969],accel_mss,speed_ms,blend_radius_m)
  movec([0.383380, -1.174583, -2.688341, -0.849465, 1.570796, 1.954177],[0.381579, -1.175976, -2.687715, -0.848698, 1.570796, 1.952375],accel_mss,speed_ms,blend_radius_m)
  movec([0.380024, -1.177137, -2.687191, -0.848061, 1.570796, 1.950821],[0.378458, -1.178259, -2.686684, -0.847446, 1.570796, 1.949255],accel_mss,speed_ms,blend_radius_m)
  movec([0.377805, -1.178710, -2.686480, -0.847199, 1.570796, 1.948602],[0.377150, -1.179149, -2.686281, -0.846959, 1.570796, 1.947946],accel_mss,speed_ms,blend_radius_m)
  movel([0.376633, -1.179481, -2.686130, -0.846778, 1.570796, 1.947430],accel_mss,speed_ms,0,blend_radius_m)
  movec([0.375988, -1.179874, -2.685951, -0.846564, 1.570796, 1.946784],[0.375339, -1.180240, -2.685785, -0.846364, 1.570796, 1.946135],accel_mss,speed_ms,blend_radius_m)
  movec([0.374616, -1.180610, -2.685617, -0.846163, 1.570796, 1.945413],[0.373895, -1.180929, -2.685471, -0.845989, 1.570796, 1.944691],accel_mss,speed_ms,blend_radius_m)
  movel([0.372745, -1.181288, -2.685308, -0.845794, 1.570796, 1.943541],accel_mss,speed_ms,0,blend_radius_m)
  movel([0.371824, -1.181368, -2.685271, -0.845750, 1.570796, 1.942620],accel_mss,speed_ms,0,blend_radius_m)
  movec([0.371263, -1.181260, -2.685320, -0.845809, 1.570796, 1.942059],[0.370806, -1.181007, -2.685436, -0.845946, 1.570796, 1.941602],accel_mss,speed_ms,blend_radius_m)
  movec([0.370459, -1.180627, -2.685609, -0.846153, 1.570796, 1.941255],[0.370230, -1.180143, -2.685829, -0.846417, 1.570796, 1.941026],accel_mss,speed_ms,blend_radius_m)
  movel([0.370158, -1.179173, -2.686270, -0.846946, 1.570796, 1.940954],accel_mss,speed_ms,0,blend_radius_m)
  movel([0.370349, -1.178357, -2.686640, -0.847392, 1.570796, 1.941145],accel_mss,speed_ms,0,blend_radius_m)
  movel([0.370830, -1.177273, -2.687130, -0.847986, 1.570796, 1.941626],accel_mss,speed_ms,0,blend_radius_m)
  movel([0.371354, -1.176395, -2.687526, -0.848468, 1.570796, 1.942150],accel_mss,speed_ms,0,blend_radius_m)
  movel([0.372210, -1.175205, -2.688062, -0.849122, 1.570796, 1.943006],accel_mss,speed_ms,0,blend_radius_m)
  movec([0.372855, -1.174408, -2.688420, -0.849561, 1.570796, 1.943651],[0.373529, -1.173627, -2.688770, -0.849992, 1.570796, 1.944325],accel_mss,speed_ms,blend_radius_m)
  movel([0.374560, -1.172504, -2.689273, -0.850612, 1.570796, 1.945357],accel_mss,speed_ms,0,blend_radius_m)
  movec([0.375805, -1.171209, -2.689850, -0.851329, 1.570796, 1.946601],[0.377074, -1.169934, -2.690417, -0.852038, 1.570796, 1.947870],accel_mss,speed_ms,blend_radius_m)
  movec([0.378289, -1.168750, -2.690943, -0.852697, 1.570796, 1.949086],[0.379521, -1.167579, -2.691460, -0.853350, 1.570796, 1.950317],accel_mss,speed_ms,blend_radius_m)
  movec([0.381418, -1.165813, -2.692239, -0.854337, 1.570796, 1.952214],[0.383338, -1.164066, -2.693005, -0.855318, 1.570796, 1.954134],accel_mss,speed_ms,blend_radius_m)
  movec([0.385625, -1.162028, -2.693896, -0.856465, 1.570796, 1.956422],[0.387934, -1.160007, -2.694775, -0.857607, 1.570796, 1.958731],accel_mss,speed_ms,blend_radius_m)
  movel([0.389088, -1.159010, -2.695207, -0.858172, 1.570796, 1.959885],accel_mss,speed_ms,0,blend_radius_m)
  movec([0.390425, -1.157864, -2.695702, -0.858823, 1.570796, 1.961222],[0.391769, -1.156723, -2.696194, -0.859472, 1.570796, 1.962566],accel_mss,speed_ms,blend_radius_m)
  movec([0.393845, -1.154988, -2.696939, -0.860462, 1.570796, 1.964642],[0.395939, -1.153272, -2.697673, -0.861443, 1.570796, 1.966736],accel_mss,speed_ms,blend_radius_m)
  movec([0.397784, -1.151798, -2.698302, -0.862289, 1.570796, 1.968581],[0.399648, -1.150354, -2.698915, -0.863120, 1.570796, 1.970444],accel_mss,speed_ms,blend_radius_m)
  movec([0.401258, -1.149148, -2.699426, -0.863815, 1.570796, 1.972055],[0.402885, -1.147981, -2.699919, -0.864490, 1.570796, 1.973681],accel_mss,speed_ms,blend_radius_m)
  speed_ms = 0.003
  movel([0.402885, -1.140599, -2.696125, -0.875666, 1.570796, 1.973681],accel_mss,speed_ms,0,blend_radius_m)
  speed_ms = 0.05
  movel([0.402885, -1.112693, -2.680709, -0.918987, 1.570796, 1.973681],accel_mss,speed_ms,0,blend_radius_m)
  #M_RunCode9
  movel([0.407472, -1.105727, -2.683497, -0.923164, 1.570796, 1.978268],accel_mss,speed_ms,0,blend_radius_m)
  #M_RunCode3
  movel([0.407472, -1.133651, -2.699003, -0.879735, 1.570796, 1.978268],accel_mss,speed_ms,0,blend_radius_m)
  speed_ms = 0.003
  movel([0.407472, -1.141043, -2.702820, -0.868526, 1.570796, 1.978268],accel_mss,speed_ms,0,blend_radius_m)
  speed_ms = 0.007
  movec([0.408985, -1.141586, -2.702595, -0.868208, 1.570796, 1.979782],[0.410294, -1.142393, -2.702259, -0.867737, 1.570796, 1.981090],accel_mss,speed_ms,blend_radius_m)
  movec([0.411019, -1.143038, -2.701991, -0.867360, 1.570796, 1.981815],[0.411654, -1.143773, -2.701684, -0.866932, 1.570796, 1.982450],accel_mss,speed_ms,blend_radius_m)
  movec([0.412395, -1.144946, -2.701194, -0.866249, 1.570796, 1.983192],[0.412961, -1.146262, -2.700642, -0.865485, 1.570796, 1.983758],accel_mss,speed_ms,blend_radius_m)
  movec([0.413256, -1.147318, -2.700198, -0.864873, 1.570796, 1.984052],[0.413437, -1.148447, -2.699722, -0.864220, 1.570796, 1.984234],accel_mss,speed_ms,blend_radius_m)
  movec([0.413503, -1.149750, -2.699171, -0.863468, 1.570796, 1.984300],[0.413429, -1.151122, -2.698589, -0.862678, 1.570796, 1.984225],accel_mss,speed_ms,blend_radius_m)
  movec([0.413322, -1.151959, -2.698233, -0.862197, 1.570796, 1.984118],[0.413168, -1.152812, -2.697870, -0.861707, 1.570796, 1.983965],accel_mss,speed_ms,blend_radius_m)
  movec([0.412886, -1.153985, -2.697369, -0.861035, 1.570796, 1.983682],[0.412515, -1.155178, -2.696858, -0.860353, 1.570796, 1.983311],accel_mss,speed_ms,blend_radius_m)
  movec([0.411879, -1.156817, -2.696153, -0.859418, 1.570796, 1.982676],[0.411107, -1.158463, -2.695443, -0.858483, 1.570796, 1.981903],accel_mss,speed_ms,blend_radius_m)
  movec([0.410259, -1.160021, -2.694769, -0.857600, 1.570796, 1.981055],[0.409317, -1.161562, -2.694099, -0.856728, 1.570796, 1.980114],accel_mss,speed_ms,blend_radius_m)
  movec([0.408751, -1.162421, -2.693725, -0.856244, 1.570796, 1.979547],[0.408162, -1.163272, -2.693353, -0.855764, 1.570796, 1.978958],accel_mss,speed_ms,blend_radius_m)
  movec([0.407339, -1.164395, -2.692861, -0.855133, 1.570796, 1.978136],[0.406478, -1.165499, -2.692376, -0.854513, 1.570796, 1.977274],accel_mss,speed_ms,blend_radius_m)
  movec([0.404894, -1.167378, -2.691549, -0.853462, 1.570796, 1.975690],[0.403227, -1.169190, -2.690747, -0.852452, 1.570796, 1.974023],accel_mss,speed_ms,blend_radius_m)
  movec([0.401709, -1.170722, -2.690067, -0.851600, 1.570796, 1.972505],[0.400150, -1.172202, -2.689407, -0.850780, 1.570796, 1.970946],accel_mss,speed_ms,blend_radius_m)
  movec([0.397468, -1.174568, -2.688348, -0.849473, 1.570796, 1.968264],[0.394717, -1.176797, -2.687345, -0.848247, 1.570796, 1.965514],accel_mss,speed_ms,blend_radius_m)
  movec([0.392783, -1.178242, -2.686692, -0.847455, 1.570796, 1.963580],[0.390822, -1.179598, -2.686077, -0.846714, 1.570796, 1.961618],accel_mss,speed_ms,blend_radius_m)
  movec([0.388916, -1.180797, -2.685531, -0.846061, 1.570796, 1.959712],[0.386995, -1.181880, -2.685037, -0.845471, 1.570796, 1.957791],accel_mss,speed_ms,blend_radius_m)
  movec([0.386035, -1.182373, -2.684812, -0.845204, 1.570796, 1.956831],[0.385075, -1.182827, -2.684604, -0.844957, 1.570796, 1.955871],accel_mss,speed_ms,blend_radius_m)
  movec([0.383264, -1.183589, -2.684255, -0.844544, 1.570796, 1.954060],[0.381470, -1.184218, -2.683967, -0.844204, 1.570796, 1.952266],accel_mss,speed_ms,blend_radius_m)
  movec([0.379623, -1.184708, -2.683742, -0.843939, 1.570796, 1.950420],[0.377838, -1.184997, -2.683609, -0.843783, 1.570796, 1.948634],accel_mss,speed_ms,blend_radius_m)
  movec([0.376588, -1.185070, -2.683575, -0.843743, 1.570796, 1.947384],[0.375396, -1.185022, -2.683597, -0.843770, 1.570796, 1.946193],accel_mss,speed_ms,blend_radius_m)
  movec([0.374712, -1.184935, -2.683637, -0.843817, 1.570796, 1.945508],[0.374052, -1.184807, -2.683696, -0.843886, 1.570796, 1.944848],accel_mss,speed_ms,blend_radius_m)
  movec([0.372577, -1.184327, -2.683917, -0.844145, 1.570796, 1.943373],[0.371284, -1.183607, -2.684247, -0.844535, 1.570796, 1.942080],accel_mss,speed_ms,blend_radius_m)
  movec([0.370602, -1.183068, -2.684494, -0.844827, 1.570796, 1.941399],[0.369993, -1.182453, -2.684776, -0.845161, 1.570796, 1.940790],accel_mss,speed_ms,blend_radius_m)
  movec([0.369652, -1.182039, -2.684965, -0.845385, 1.570796, 1.940449],[0.369338, -1.181600, -2.685165, -0.845624, 1.570796, 1.940135],accel_mss,speed_ms,blend_radius_m)
  movec([0.368757, -1.180580, -2.685630, -0.846179, 1.570796, 1.939553],[0.368307, -1.179455, -2.686141, -0.846792, 1.570796, 1.939103],accel_mss,speed_ms,blend_radius_m)
  movec([0.367915, -1.177606, -2.686980, -0.847804, 1.570796, 1.938712],[0.367876, -1.175551, -2.687906, -0.848931, 1.570796, 1.938672],accel_mss,speed_ms,blend_radius_m)
  movec([0.367946, -1.174773, -2.688256, -0.849360, 1.570796, 1.938743],[0.368060, -1.173976, -2.688614, -0.849799, 1.570796, 1.938857],accel_mss,speed_ms,blend_radius_m)
  movec([0.368294, -1.172843, -2.689121, -0.850425, 1.570796, 1.939090],[0.368615, -1.171684, -2.689638, -0.851066, 1.570796, 1.939411],accel_mss,speed_ms,blend_radius_m)
  movec([0.369182, -1.170088, -2.690349, -0.851952, 1.570796, 1.939979],[0.369895, -1.168473, -2.691065, -0.852851, 1.570796, 1.940691],accel_mss,speed_ms,blend_radius_m)
  movec([0.370684, -1.166934, -2.691745, -0.853710, 1.570796, 1.941481],[0.371573, -1.165400, -2.692420, -0.854569, 1.570796, 1.942369],accel_mss,speed_ms,blend_radius_m)
  movec([0.372113, -1.164540, -2.692798, -0.855051, 1.570796, 1.942909],[0.372677, -1.163684, -2.693173, -0.855533, 1.570796, 1.943474],accel_mss,speed_ms,blend_radius_m)
  movec([0.373473, -1.162547, -2.693669, -0.856173, 1.570796, 1.944269],[0.374311, -1.161424, -2.694159, -0.856806, 1.570796, 1.945108],accel_mss,speed_ms,blend_radius_m)
  movec([0.375865, -1.159503, -2.694993, -0.857893, 1.570796, 1.946661],[0.377516, -1.157635, -2.695801, -0.858953, 1.570796, 1.948313],accel_mss,speed_ms,blend_radius_m)
  movec([0.378917, -1.156162, -2.696435, -0.859792, 1.570796, 1.949713],[0.380363, -1.154727, -2.697051, -0.860611, 1.570796, 1.951159],accel_mss,speed_ms,blend_radius_m)
  movec([0.381583, -1.153573, -2.697545, -0.861271, 1.570796, 1.952379],[0.382825, -1.152443, -2.698027, -0.861919, 1.570796, 1.953622],accel_mss,speed_ms,blend_radius_m)
  movel([0.383626, -1.151739, -2.698327, -0.862323, 1.570796, 1.954422],accel_mss,speed_ms,0,blend_radius_m)
  movec([0.384792, -1.150742, -2.698751, -0.862896, 1.570796, 1.955588],[0.385973, -1.149766, -2.699164, -0.863459, 1.570796, 1.956769],accel_mss,speed_ms,blend_radius_m)
  movec([0.387467, -1.148589, -2.699662, -0.864138, 1.570796, 1.958264],[0.388985, -1.147460, -2.700138, -0.864791, 1.570796, 1.959781],accel_mss,speed_ms,blend_radius_m)
  movec([0.390492, -1.146408, -2.700581, -0.865400, 1.570796, 1.961288],[0.392016, -1.145417, -2.700997, -0.865975, 1.570796, 1.962812],accel_mss,speed_ms,blend_radius_m)
  movec([0.393459, -1.144550, -2.701359, -0.866479, 1.570796, 1.964256],[0.394910, -1.143753, -2.701693, -0.866943, 1.570796, 1.965707],accel_mss,speed_ms,blend_radius_m)
  movel([0.396168, -1.143129, -2.701953, -0.867307, 1.570796, 1.966964],accel_mss,speed_ms,0,blend_radius_m)
  movec([0.398061, -1.142303, -2.702297, -0.867789, 1.570796, 1.968857],[0.399936, -1.141621, -2.702581, -0.868188, 1.570796, 1.970732],accel_mss,speed_ms,blend_radius_m)
  movec([0.401835, -1.141103, -2.702795, -0.868491, 1.570796, 1.972632],[0.403666, -1.140805, -2.702919, -0.868665, 1.570796, 1.974463],accel_mss,speed_ms,blend_radius_m)
  movec([0.404803, -1.140737, -2.702947, -0.868705, 1.570796, 1.975600],[0.405889, -1.140777, -2.702931, -0.868681, 1.570796, 1.976685],accel_mss,speed_ms,blend_radius_m)
  movel([0.406217, -1.140814, -2.702915, -0.868660, 1.570796, 1.977013],accel_mss,speed_ms,0,blend_radius_m)
  movec([0.406855, -1.140911, -2.702875, -0.868603, 1.570796, 1.977651],[0.407472, -1.141043, -2.702820, -0.868526, 1.570796, 1.978268],accel_mss,speed_ms,blend_radius_m)
  speed_ms = 0.003
  movel([0.407472, -1.133651, -2.699003, -0.879735, 1.570796, 1.978268],accel_mss,speed_ms,0,blend_radius_m)
  speed_ms = 0.05
  movel([0.407472, -1.105727, -2.683497, -0.923164, 1.570796, 1.978268],accel_mss,speed_ms,0,blend_radius_m)
  #M_RunCode9
  movel([0.476572, -1.340603, -2.560956, -0.810830, 1.570796, 2.047369],accel_mss,speed_ms,0,blend_radius_m)
  #M_RunCode3
  movel([0.476572, -1.365929, -2.573377, -0.773083, 1.570796, 2.047369],accel_mss,speed_ms,0,blend_radius_m)
  speed_ms = 0.003
  movel([0.476572, -1.372510, -2.576410, -0.763468, 1.570796, 2.047369],accel_mss,speed_ms,0,blend_radius_m)
  speed_ms = 0.007
  movec([0.477638, -1.371894, -2.576838, -0.763657, 1.570796, 2.048435],[0.478730, -1.371375, -2.577198, -0.763816, 1.570796, 2.049526],accel_mss,speed_ms,blend_radius_m)
  movec([0.479616, -1.371029, -2.577437, -0.763922, 1.570796, 2.050412],[0.480501, -1.370749, -2.577631, -0.764009, 1.570796, 2.051297],accel_mss,speed_ms,blend_radius_m)
  movec([0.481091, -1.370596, -2.577737, -0.764056, 1.570796, 2.051887],[0.481676, -1.370469, -2.577825, -0.764095, 1.570796, 2.052472],accel_mss,speed_ms,blend_radius_m)
  movec([0.483374, -1.370194, -2.578015, -0.764180, 1.570796, 2.054170],[0.485035, -1.370041, -2.578121, -0.764227, 1.570796, 2.055831],accel_mss,speed_ms,blend_radius_m)
  movec([0.485983, -1.370008, -2.578144, -0.764237, 1.570796, 2.056779],[0.486913, -1.370016, -2.578138, -0.764235, 1.570796, 2.057709],accel_mss,speed_ms,blend_radius_m)
  movec([0.487413, -1.370034, -2.578126, -0.764229, 1.570796, 2.058210],[0.487911, -1.370057, -2.578110, -0.764222, 1.570796, 2.058707],accel_mss,speed_ms,blend_radius_m)
  movec([0.489153, -1.370128, -2.578061, -0.764200, 1.570796, 2.059949],[0.490387, -1.370214, -2.578001, -0.764174, 1.570796, 2.061184],accel_mss,speed_ms,blend_radius_m)
  movec([0.491956, -1.370346, -2.577910, -0.764133, 1.570796, 2.062753],[0.493517, -1.370492, -2.577809, -0.764088, 1.570796, 2.064313],accel_mss,speed_ms,blend_radius_m)
  movec([0.495586, -1.370710, -2.577658, -0.764021, 1.570796, 2.066383],[0.497669, -1.370902, -2.577525, -0.763962, 1.570796, 2.068466],accel_mss,speed_ms,blend_radius_m)
  movec([0.498437, -1.370962, -2.577484, -0.763943, 1.570796, 2.069234],[0.499210, -1.371013, -2.577449, -0.763927, 1.570796, 2.070007],accel_mss,speed_ms,blend_radius_m)
  movel([0.499591, -1.371034, -2.577434, -0.763921, 1.570796, 2.070387],accel_mss,speed_ms,0,blend_radius_m)
  movec([0.500908, -1.371058, -2.577418, -0.763914, 1.570796, 2.071705],[0.502261, -1.370999, -2.577458, -0.763932, 1.570796, 2.073057],accel_mss,speed_ms,blend_radius_m)
  movec([0.503311, -1.370895, -2.577530, -0.763964, 1.570796, 2.074108],[0.504378, -1.370738, -2.577639, -0.764012, 1.570796, 2.075175],accel_mss,speed_ms,blend_radius_m)
  movec([0.505276, -1.370551, -2.577768, -0.764070, 1.570796, 2.076073],[0.506186, -1.370295, -2.577945, -0.764149, 1.570796, 2.076982],accel_mss,speed_ms,blend_radius_m)
  movec([0.506990, -1.370008, -2.578143, -0.764237, 1.570796, 2.077787],[0.507792, -1.369657, -2.578386, -0.764346, 1.570796, 2.078588],accel_mss,speed_ms,blend_radius_m)
  movec([0.508324, -1.369386, -2.578573, -0.764430, 1.570796, 2.079120],[0.508848, -1.369088, -2.578779, -0.764522, 1.570796, 2.079645],accel_mss,speed_ms,blend_radius_m)
  movec([0.509372, -1.368759, -2.579006, -0.764625, 1.570796, 2.080168],[0.509886, -1.368408, -2.579248, -0.764734, 1.570796, 2.080682],accel_mss,speed_ms,blend_radius_m)
  movel([0.510708, -1.367767, -2.579688, -0.764933, 1.570796, 2.081505],accel_mss,speed_ms,0,blend_radius_m)
  movel([0.511486, -1.367035, -2.580192, -0.765162, 1.570796, 2.082282],accel_mss,speed_ms,0,blend_radius_m)
  movel([0.512101, -1.366307, -2.580691, -0.765391, 1.570796, 2.082898],accel_mss,speed_ms,0,blend_radius_m)
  movel([0.512527, -1.365658, -2.581136, -0.765595, 1.570796, 2.083324],accel_mss,speed_ms,0,blend_radius_m)
  movel([0.512670, -1.365398, -2.581314, -0.765677, 1.570796, 2.083466],accel_mss,speed_ms,0,blend_radius_m)
  movec([0.512915, -1.364868, -2.581677, -0.765844, 1.570796, 2.083712],[0.513109, -1.364339, -2.582038, -0.766012, 1.570796, 2.083906],accel_mss,speed_ms,blend_radius_m)
  movec([0.513296, -1.363497, -2.582613, -0.766279, 1.570796, 2.084092],[0.513307, -1.362704, -2.583153, -0.766532, 1.570796, 2.084103],accel_mss,speed_ms,blend_radius_m)
  movel([0.513144, -1.361959, -2.583659, -0.766770, 1.570796, 2.083941],accel_mss,speed_ms,0,blend_radius_m)
  movec([0.512991, -1.361593, -2.583908, -0.766888, 1.570796, 2.083788],[0.512798, -1.361253, -2.584139, -0.766997, 1.570796, 2.083594],accel_mss,speed_ms,blend_radius_m)
  movel([0.512404, -1.360812, -2.584438, -0.767139, 1.570796, 2.083201],accel_mss,speed_ms,0,blend_radius_m)
  movel([0.512096, -1.360618, -2.584569, -0.767201, 1.570796, 2.082893],accel_mss,speed_ms,0,blend_radius_m)
  movel([0.511903, -1.360543, -2.584620, -0.767225, 1.570796, 2.082700],accel_mss,speed_ms,0,blend_radius_m)
  movel([0.511407, -1.360467, -2.584672, -0.767250, 1.570796, 2.082203],accel_mss,speed_ms,0,blend_radius_m)
  movel([0.510990, -1.360509, -2.584643, -0.767237, 1.570796, 2.081787],accel_mss,speed_ms,0,blend_radius_m)
  movel([0.510805, -1.360560, -2.584609, -0.767220, 1.570796, 2.081601],accel_mss,speed_ms,0,blend_radius_m)
  movel([0.510542, -1.360664, -2.584539, -0.767187, 1.570796, 2.081338],accel_mss,speed_ms,0,blend_radius_m)
  movel([0.510272, -1.360810, -2.584439, -0.767139, 1.570796, 2.081068],accel_mss,speed_ms,0,blend_radius_m)
  movel([0.510129, -1.360910, -2.584372, -0.767107, 1.570796, 2.080925],accel_mss,speed_ms,0,blend_radius_m)
  movel([0.509789, -1.361222, -2.584160, -0.767007, 1.570796, 2.080586],accel_mss,speed_ms,0,blend_radius_m)
  movel([0.509406, -1.361672, -2.583854, -0.766862, 1.570796, 2.080203],accel_mss,speed_ms,0,blend_radius_m)
  movel([0.509276, -1.361844, -2.583738, -0.766807, 1.570796, 2.080073],accel_mss,speed_ms,0,blend_radius_m)
  movel([0.508726, -1.362523, -2.583276, -0.766590, 1.570796, 2.079523],accel_mss,speed_ms,0,blend_radius_m)
  movel([0.508365, -1.362908, -2.583014, -0.766467, 1.570796, 2.079161],accel_mss,speed_ms,0,blend_radius_m)
  movel([0.508114, -1.363139, -2.582856, -0.766393, 1.570796, 2.078910],accel_mss,speed_ms,0,blend_radius_m)
  movel([0.507504, -1.363602, -2.582541, -0.766246, 1.570796, 2.078300],accel_mss,speed_ms,0,blend_radius_m)
  movel([0.506658, -1.364125, -2.582184, -0.766080, 1.570796, 2.077454],accel_mss,speed_ms,0,blend_radius_m)
  movel([0.505674, -1.364573, -2.581878, -0.765938, 1.570796, 2.076471],accel_mss,speed_ms,0,blend_radius_m)
  movel([0.504957, -1.364769, -2.581744, -0.765876, 1.570796, 2.075753],accel_mss,speed_ms,0,blend_radius_m)
  movel([0.504249, -1.364826, -2.581705, -0.765858, 1.570796, 2.075045],accel_mss,speed_ms,0,blend_radius_m)
  movel([0.503700, -1.364758, -2.581752, -0.765879, 1.570796, 2.074497],accel_mss,speed_ms,0,blend_radius_m)
  movel([0.503226, -1.364612, -2.581851, -0.765925, 1.570796, 2.074023],accel_mss,speed_ms,0,blend_radius_m)
  movec([0.502704, -1.364341, -2.582036, -0.766011, 1.570796, 2.073500],[0.502273, -1.363975, -2.582286, -0.766127, 1.570796, 2.073069],accel_mss,speed_ms,blend_radius_m)
  movec([0.502000, -1.363627, -2.582524, -0.766238, 1.570796, 2.072796],[0.501783, -1.363237, -2.582790, -0.766362, 1.570796, 2.072579],accel_mss,speed_ms,blend_radius_m)
  movel([0.501720, -1.363091, -2.582890, -0.766409, 1.570796, 2.072516],accel_mss,speed_ms,0,blend_radius_m)
  movec([0.501586, -1.362683, -2.583167, -0.766539, 1.570796, 2.072383],[0.501502, -1.362248, -2.583463, -0.766678, 1.570796, 2.072298],accel_mss,speed_ms,blend_radius_m)
  movec([0.501476, -1.361808, -2.583762, -0.766819, 1.570796, 2.072272],[0.501509, -1.361346, -2.584076, -0.766967, 1.570796, 2.072305],accel_mss,speed_ms,blend_radius_m)
  movel([0.501664, -1.360624, -2.584566, -0.767200, 1.570796, 2.072461],accel_mss,speed_ms,0,blend_radius_m)
  movel([0.501832, -1.360146, -2.584889, -0.767354, 1.570796, 2.072628],accel_mss,speed_ms,0,blend_radius_m)
  movel([0.502094, -1.359605, -2.585255, -0.767529, 1.570796, 2.072891],accel_mss,speed_ms,0,blend_radius_m)
  movec([0.502484, -1.359018, -2.585652, -0.767719, 1.570796, 2.073280],[0.502969, -1.358465, -2.586025, -0.767898, 1.570796, 2.073765],accel_mss,speed_ms,blend_radius_m)
  movel([0.503683, -1.357843, -2.586445, -0.768101, 1.570796, 2.074480],accel_mss,speed_ms,0,blend_radius_m)
  movel([0.504261, -1.357440, -2.586717, -0.768233, 1.570796, 2.075057],accel_mss,speed_ms,0,blend_radius_m)
  movel([0.504501, -1.357290, -2.586817, -0.768282, 1.570796, 2.075297],accel_mss,speed_ms,0,blend_radius_m)
  movec([0.505038, -1.356989, -2.587020, -0.768380, 1.570796, 2.075834],[0.505584, -1.356726, -2.587197, -0.768466, 1.570796, 2.076380],accel_mss,speed_ms,blend_radius_m)
  movel([0.506450, -1.356404, -2.587413, -0.768572, 1.570796, 2.077247],accel_mss,speed_ms,0,blend_radius_m)
  movec([0.507086, -1.356248, -2.587518, -0.768623, 1.570796, 2.077882],[0.507704, -1.356166, -2.587573, -0.768650, 1.570796, 2.078500],accel_mss,speed_ms,blend_radius_m)
  movec([0.508259, -1.356155, -2.587581, -0.768654, 1.570796, 2.079055],[0.508785, -1.356203, -2.587548, -0.768638, 1.570796, 2.079581],accel_mss,speed_ms,blend_radius_m)
  movel([0.509584, -1.356391, -2.587422, -0.768576, 1.570796, 2.080380],accel_mss,speed_ms,0,blend_radius_m)
  movel([0.510167, -1.356624, -2.587265, -0.768500, 1.570796, 2.080963],accel_mss,speed_ms,0,blend_radius_m)
  movec([0.510642, -1.356874, -2.587097, -0.768418, 1.570796, 2.081439],[0.511085, -1.357160, -2.586905, -0.768324, 1.570796, 2.081882],accel_mss,speed_ms,blend_radius_m)
  movec([0.511789, -1.357728, -2.586523, -0.768139, 1.570796, 2.082585],[0.512408, -1.358372, -2.586088, -0.767929, 1.570796, 2.083204],accel_mss,speed_ms,blend_radius_m)
  movec([0.512892, -1.359008, -2.585659, -0.767722, 1.570796, 2.083688],[0.513315, -1.359688, -2.585199, -0.767502, 1.570796, 2.084111],accel_mss,speed_ms,blend_radius_m)
  movec([0.513703, -1.360440, -2.584690, -0.767259, 1.570796, 2.084499],[0.514040, -1.361223, -2.584159, -0.767007, 1.570796, 2.084836],accel_mss,speed_ms,blend_radius_m)
  movec([0.514358, -1.362132, -2.583542, -0.766715, 1.570796, 2.085154],[0.514618, -1.363073, -2.582902, -0.766414, 1.570796, 2.085414],accel_mss,speed_ms,blend_radius_m)
  movec([0.514878, -1.364458, -2.581957, -0.765974, 1.570796, 2.085675],[0.515004, -1.365903, -2.580968, -0.765518, 1.570796, 2.085800],accel_mss,speed_ms,blend_radius_m)
  movec([0.514996, -1.367190, -2.580085, -0.765114, 1.570796, 2.085792],[0.514872, -1.368513, -2.579175, -0.764701, 1.570796, 2.085668],accel_mss,speed_ms,blend_radius_m)
  movec([0.514746, -1.369308, -2.578627, -0.764454, 1.570796, 2.085543],[0.514582, -1.370113, -2.578071, -0.764205, 1.570796, 2.085378],accel_mss,speed_ms,blend_radius_m)
  movec([0.514393, -1.370810, -2.577589, -0.763990, 1.570796, 2.085189],[0.514144, -1.371514, -2.577101, -0.763773, 1.570796, 2.084940],accel_mss,speed_ms,blend_radius_m)
  movec([0.513836, -1.372214, -2.576616, -0.763559, 1.570796, 2.084632],[0.513463, -1.372910, -2.576133, -0.763347, 1.570796, 2.084259],accel_mss,speed_ms,blend_radius_m)
  movec([0.512833, -1.373863, -2.575470, -0.763057, 1.570796, 2.083629],[0.512088, -1.374776, -2.574833, -0.762780, 1.570796, 2.082884],accel_mss,speed_ms,blend_radius_m)
  movec([0.511416, -1.375473, -2.574346, -0.762570, 1.570796, 2.082212],[0.510693, -1.376128, -2.573888, -0.762373, 1.570796, 2.081489],accel_mss,speed_ms,blend_radius_m)
  movec([0.510005, -1.376682, -2.573500, -0.762206, 1.570796, 2.080802],[0.509293, -1.377201, -2.573136, -0.762051, 1.570796, 2.080089],accel_mss,speed_ms,blend_radius_m)
  movec([0.508426, -1.377772, -2.572736, -0.761881, 1.570796, 2.079223],[0.507541, -1.378296, -2.572368, -0.761725, 1.570796, 2.078337],accel_mss,speed_ms,blend_radius_m)
  movec([0.506678, -1.378750, -2.572049, -0.761590, 1.570796, 2.077474],[0.505805, -1.379151, -2.571767, -0.761471, 1.570796, 2.076601],accel_mss,speed_ms,blend_radius_m)
  movec([0.504862, -1.379515, -2.571510, -0.761364, 1.570796, 2.075658],[0.503921, -1.379806, -2.571305, -0.761278, 1.570796, 2.074718],accel_mss,speed_ms,blend_radius_m)
  movel([0.503331, -1.379954, -2.571201, -0.761234, 1.570796, 2.074128],accel_mss,speed_ms,0,blend_radius_m)
  movec([0.502204, -1.380177, -2.571043, -0.761168, 1.570796, 2.073000],[0.501093, -1.380336, -2.570931, -0.761121, 1.570796, 2.071889],accel_mss,speed_ms,blend_radius_m)
  movec([0.499968, -1.380433, -2.570863, -0.761093, 1.570796, 2.070764],[0.498870, -1.380457, -2.570846, -0.761086, 1.570796, 2.069667],accel_mss,speed_ms,blend_radius_m)
  movel([0.498028, -1.380434, -2.570862, -0.761093, 1.570796, 2.068824],accel_mss,speed_ms,0,blend_radius_m)
  movec([0.497047, -1.380386, -2.570896, -0.761107, 1.570796, 2.067844],[0.496076, -1.380319, -2.570943, -0.761127, 1.570796, 2.066873],accel_mss,speed_ms,blend_radius_m)
  movec([0.494926, -1.380217, -2.571015, -0.761156, 1.570796, 2.065722],[0.493785, -1.380099, -2.571099, -0.761191, 1.570796, 2.064581],accel_mss,speed_ms,blend_radius_m)
  movec([0.492168, -1.379960, -2.571196, -0.761232, 1.570796, 2.062965],[0.490534, -1.379857, -2.571269, -0.761263, 1.570796, 2.061330],accel_mss,speed_ms,blend_radius_m)
  movec([0.489903, -1.379830, -2.571288, -0.761271, 1.570796, 2.060699],[0.489267, -1.379814, -2.571300, -0.761275, 1.570796, 2.060064],accel_mss,speed_ms,blend_radius_m)
  movel([0.488955, -1.379811, -2.571302, -0.761276, 1.570796, 2.059751],accel_mss,speed_ms,0,blend_radius_m)
  movec([0.488309, -1.379821, -2.571295, -0.761273, 1.570796, 2.059106],[0.487654, -1.379857, -2.571270, -0.761263, 1.570796, 2.058450],accel_mss,speed_ms,blend_radius_m)
  movec([0.486783, -1.379946, -2.571206, -0.761236, 1.570796, 2.057579],[0.485898, -1.380084, -2.571109, -0.761196, 1.570796, 2.056695],accel_mss,speed_ms,blend_radius_m)
  movel([0.484912, -1.380287, -2.570966, -0.761136, 1.570796, 2.055708],accel_mss,speed_ms,0,blend_radius_m)
  movel([0.483968, -1.380547, -2.570783, -0.761060, 1.570796, 2.054764],accel_mss,speed_ms,0,blend_radius_m)
  movec([0.482894, -1.380941, -2.570504, -0.760944, 1.570796, 2.053691],[0.481830, -1.381439, -2.570152, -0.760798, 1.570796, 2.052626],accel_mss,speed_ms,blend_radius_m)
  movec([0.481307, -1.381724, -2.569951, -0.760714, 1.570796, 2.052104],[0.480793, -1.382032, -2.569733, -0.760625, 1.570796, 2.051589],accel_mss,speed_ms,blend_radius_m)
  movel([0.481119, -1.382775, -2.569206, -0.760408, 1.570796, 2.051915],accel_mss,speed_ms,0,blend_radius_m)
  movec([0.481572, -1.383717, -2.568537, -0.760135, 1.570796, 2.052368],[0.482086, -1.384619, -2.567896, -0.759874, 1.570796, 2.052882],accel_mss,speed_ms,blend_radius_m)
  movec([0.482531, -1.385280, -2.567425, -0.759684, 1.570796, 2.053327],[0.483025, -1.385903, -2.566981, -0.759506, 1.570796, 2.053822],accel_mss,speed_ms,blend_radius_m)
  movec([0.483426, -1.386334, -2.566673, -0.759382, 1.570796, 2.054222],[0.483860, -1.386736, -2.566386, -0.759268, 1.570796, 2.054656],accel_mss,speed_ms,blend_radius_m)
  movec([0.484286, -1.387076, -2.566142, -0.759171, 1.570796, 2.055083],[0.484743, -1.387386, -2.565920, -0.759082, 1.570796, 2.055540],accel_mss,speed_ms,blend_radius_m)
  movec([0.485234, -1.387660, -2.565724, -0.759005, 1.570796, 2.056030],[0.485759, -1.387894, -2.565557, -0.758938, 1.570796, 2.056555],accel_mss,speed_ms,blend_radius_m)
  movel([0.486303, -1.388081, -2.565422, -0.758885, 1.570796, 2.057100],accel_mss,speed_ms,0,blend_radius_m)
  movec([0.487020, -1.388255, -2.565298, -0.758836, 1.570796, 2.057817],[0.487775, -1.388369, -2.565216, -0.758804, 1.570796, 2.058572],accel_mss,speed_ms,blend_radius_m)
  movec([0.488558, -1.388417, -2.565181, -0.758790, 1.570796, 2.059354],[0.489372, -1.388396, -2.565197, -0.758796, 1.570796, 2.060168],accel_mss,speed_ms,blend_radius_m)
  movec([0.490575, -1.388239, -2.565309, -0.758841, 1.570796, 2.061372],[0.491813, -1.387936, -2.565527, -0.758927, 1.570796, 2.062609],accel_mss,speed_ms,blend_radius_m)
  movec([0.492670, -1.387648, -2.565733, -0.759008, 1.570796, 2.063466],[0.493526, -1.387302, -2.565981, -0.759106, 1.570796, 2.064322],accel_mss,speed_ms,blend_radius_m)
  movel([0.484370, -1.392896, -2.561954, -0.757539, 1.570796, 2.055166],accel_mss,speed_ms,0,blend_radius_m)
  movel([0.475642, -1.373100, -2.576000, -0.763289, 1.570796, 2.046438],accel_mss,speed_ms,0,blend_radius_m)
  movel([0.476572, -1.372510, -2.576410, -0.763468, 1.570796, 2.047369],accel_mss,speed_ms,0,blend_radius_m)
  speed_ms = 0.003
  movel([0.476572, -1.365929, -2.573377, -0.773083, 1.570796, 2.047369],accel_mss,speed_ms,0,blend_radius_m)
  speed_ms = 0.05
  movel([0.476572, -1.340603, -2.560956, -0.810830, 1.570796, 2.047369],accel_mss,speed_ms,0,blend_radius_m)
  #M_RunCode9
  movel([0.490591, -1.360792, -2.547307, -0.804290, 1.570796, 2.061387],accel_mss,speed_ms,0,blend_radius_m)
  #M_RunCode3
  movel([0.490591, -1.385747, -2.559471, -0.767170, 1.570796, 2.061387],accel_mss,speed_ms,0,blend_radius_m)
  speed_ms = 0.003
  movel([0.490591, -1.392225, -2.562440, -0.757725, 1.570796, 2.061387],accel_mss,speed_ms,0,blend_radius_m)
  speed_ms = 0.007
  movel([0.491526, -1.391640, -2.562862, -0.757887, 1.570796, 2.062323],accel_mss,speed_ms,0,blend_radius_m)
  movel([0.492329, -1.391273, -2.563127, -0.757989, 1.570796, 2.063125],accel_mss,speed_ms,0,blend_radius_m)
  movel([0.493004, -1.391076, -2.563269, -0.758044, 1.570796, 2.063800],accel_mss,speed_ms,0,blend_radius_m)
  movel([0.493870, -1.390998, -2.563325, -0.758066, 1.570796, 2.064667],accel_mss,speed_ms,0,blend_radius_m)
  movel([0.494372, -1.391061, -2.563280, -0.758048, 1.570796, 2.065168],accel_mss,speed_ms,0,blend_radius_m)
  movel([0.494838, -1.391195, -2.563183, -0.758011, 1.570796, 2.065634],accel_mss,speed_ms,0,blend_radius_m)
  movec([0.495332, -1.391439, -2.563007, -0.757943, 1.570796, 2.066128],[0.495743, -1.391769, -2.562769, -0.757851, 1.570796, 2.066539],accel_mss,speed_ms,blend_radius_m)
  movec([0.495989, -1.392056, -2.562562, -0.757772, 1.570796, 2.066785],[0.496191, -1.392376, -2.562330, -0.757683, 1.570796, 2.066987],accel_mss,speed_ms,blend_radius_m)
  movec([0.496383, -1.392821, -2.562009, -0.757560, 1.570796, 2.067179],[0.496506, -1.393304, -2.561659, -0.757427, 1.570796, 2.067303],accel_mss,speed_ms,blend_radius_m)
  movel([0.496545, -1.394073, -2.561101, -0.757215, 1.570796, 2.067341],accel_mss,speed_ms,0,blend_radius_m)
  movec([0.496490, -1.394505, -2.560788, -0.757097, 1.570796, 2.067287],[0.496383, -1.394948, -2.560466, -0.756975, 1.570796, 2.067180],accel_mss,speed_ms,blend_radius_m)
  movel([0.496196, -1.395467, -2.560088, -0.756834, 1.570796, 2.066993],accel_mss,speed_ms,0,blend_radius_m)
  movel([0.495909, -1.396039, -2.559672, -0.756678, 1.570796, 2.066705],accel_mss,speed_ms,0,blend_radius_m)
  movec([0.495521, -1.396596, -2.559266, -0.756527, 1.570796, 2.066317],[0.495042, -1.397114, -2.558887, -0.756387, 1.570796, 2.065839],accel_mss,speed_ms,blend_radius_m)
  movec([0.494595, -1.397506, -2.558602, -0.756282, 1.570796, 2.065392],[0.494115, -1.397857, -2.558345, -0.756187, 1.570796, 2.064911],accel_mss,speed_ms,blend_radius_m)
  movec([0.493614, -1.398172, -2.558115, -0.756102, 1.570796, 2.064410],[0.493101, -1.398453, -2.557909, -0.756027, 1.570796, 2.063897],accel_mss,speed_ms,blend_radius_m)
  movel([0.492578, -1.398687, -2.557737, -0.755964, 1.570796, 2.063374],accel_mss,speed_ms,0,blend_radius_m)
  movel([0.492315, -1.398777, -2.557672, -0.755940, 1.570796, 2.063111],accel_mss,speed_ms,0,blend_radius_m)
  movel([0.491822, -1.398899, -2.557583, -0.755908, 1.570796, 2.062618],accel_mss,speed_ms,0,blend_radius_m)
  movel([0.491133, -1.399006, -2.557504, -0.755879, 1.570796, 2.061929],accel_mss,speed_ms,0,blend_radius_m)
  movel([0.490570, -1.399094, -2.557439, -0.755855, 1.570796, 2.061366],accel_mss,speed_ms,0,blend_radius_m)
  movel([0.490111, -1.399233, -2.557337, -0.755818, 1.570796, 2.060907],accel_mss,speed_ms,0,blend_radius_m)
  movel([0.489917, -1.399332, -2.557265, -0.755792, 1.570796, 2.060713],accel_mss,speed_ms,0,blend_radius_m)
  movel([0.489782, -1.399419, -2.557201, -0.755769, 1.570796, 2.060579],accel_mss,speed_ms,0,blend_radius_m)
  movel([0.489571, -1.399580, -2.557083, -0.755726, 1.570796, 2.060367],accel_mss,speed_ms,0,blend_radius_m)
  movel([0.489215, -1.399960, -2.556804, -0.755625, 1.570796, 2.060011],accel_mss,speed_ms,0,blend_radius_m)
  movel([0.488947, -1.400410, -2.556474, -0.755505, 1.570796, 2.059744],accel_mss,speed_ms,0,blend_radius_m)
  movel([0.488832, -1.400703, -2.556258, -0.755428, 1.570796, 2.059628],accel_mss,speed_ms,0,blend_radius_m)
  movec([0.488718, -1.401176, -2.555910, -0.755303, 1.570796, 2.059514],[0.488696, -1.401627, -2.555579, -0.755184, 1.570796, 2.059492],accel_mss,speed_ms,blend_radius_m)
  movel([0.488847, -1.402325, -2.555064, -0.755000, 1.570796, 2.059643],accel_mss,speed_ms,0,blend_radius_m)
  movec([0.489073, -1.402778, -2.554730, -0.754882, 1.570796, 2.059869],[0.489363, -1.403187, -2.554428, -0.754775, 1.570796, 2.060159],accel_mss,speed_ms,blend_radius_m)
  movec([0.489983, -1.403738, -2.554020, -0.754631, 1.570796, 2.060779],[0.490772, -1.404115, -2.553741, -0.754533, 1.570796, 2.061568],accel_mss,speed_ms,blend_radius_m)
  movec([0.491256, -1.404245, -2.553645, -0.754499, 1.570796, 2.062052],[0.491770, -1.404327, -2.553584, -0.754478, 1.570796, 2.062567],accel_mss,speed_ms,blend_radius_m)
  movel([0.492428, -1.404362, -2.553558, -0.754469, 1.570796, 2.063225],accel_mss,speed_ms,0,blend_radius_m)
  movel([0.492995, -1.404343, -2.553572, -0.754474, 1.570796, 2.063792],accel_mss,speed_ms,0,blend_radius_m)
  movec([0.493581, -1.404281, -2.553618, -0.754490, 1.570796, 2.064378],[0.494179, -1.404174, -2.553697, -0.754518, 1.570796, 2.064975],accel_mss,speed_ms,blend_radius_m)
  movec([0.494856, -1.404007, -2.553821, -0.754561, 1.570796, 2.065652],[0.495537, -1.403789, -2.553982, -0.754618, 1.570796, 2.066333],accel_mss,speed_ms,blend_radius_m)
  movec([0.496279, -1.403504, -2.554193, -0.754692, 1.570796, 2.067075],[0.497017, -1.403174, -2.554437, -0.754778, 1.570796, 2.067813],accel_mss,speed_ms,blend_radius_m)
  movec([0.497953, -1.402691, -2.554794, -0.754904, 1.570796, 2.068750],[0.498873, -1.402154, -2.555190, -0.755045, 1.570796, 2.069670],accel_mss,speed_ms,blend_radius_m)
  movec([0.499614, -1.401667, -2.555549, -0.755173, 1.570796, 2.070410],[0.500331, -1.401140, -2.555937, -0.755312, 1.570796, 2.071127],accel_mss,speed_ms,blend_radius_m)
  movec([0.501425, -1.400204, -2.556625, -0.755560, 1.570796, 2.072221],[0.502414, -1.399180, -2.557377, -0.755833, 1.570796, 2.073210],accel_mss,speed_ms,blend_radius_m)
  movec([0.502887, -1.398614, -2.557791, -0.755984, 1.570796, 2.073684],[0.503328, -1.398034, -2.558216, -0.756139, 1.570796, 2.074125],accel_mss,speed_ms,blend_radius_m)
  movec([0.503654, -1.397559, -2.558563, -0.756267, 1.570796, 2.074450],[0.503951, -1.397077, -2.558915, -0.756397, 1.570796, 2.074747],accel_mss,speed_ms,blend_radius_m)
  movec([0.504394, -1.396252, -2.559516, -0.756620, 1.570796, 2.075191],[0.504762, -1.395423, -2.560120, -0.756846, 1.570796, 2.075558],accel_mss,speed_ms,blend_radius_m)
  movec([0.505074, -1.394548, -2.560756, -0.757085, 1.570796, 2.075870],[0.505313, -1.393681, -2.561386, -0.757323, 1.570796, 2.076109],accel_mss,speed_ms,blend_radius_m)
  movec([0.505470, -1.392917, -2.561939, -0.757533, 1.570796, 2.076267],[0.505582, -1.392163, -2.562484, -0.757742, 1.570796, 2.076378],accel_mss,speed_ms,blend_radius_m)
  movec([0.505635, -1.391619, -2.562877, -0.757893, 1.570796, 2.076431],[0.505663, -1.391081, -2.563265, -0.758043, 1.570796, 2.076459],accel_mss,speed_ms,blend_radius_m)
  movec([0.505649, -1.390029, -2.564023, -0.758337, 1.570796, 2.076445],[0.505554, -1.389007, -2.564758, -0.758624, 1.570796, 2.076351],accel_mss,speed_ms,blend_radius_m)
  movec([0.505375, -1.387961, -2.565509, -0.758919, 1.570796, 2.076171],[0.505123, -1.386949, -2.566233, -0.759207, 1.570796, 2.075919],accel_mss,speed_ms,blend_radius_m)
  movec([0.504850, -1.386074, -2.566858, -0.759457, 1.570796, 2.075646],[0.504535, -1.385222, -2.567466, -0.759701, 1.570796, 2.075331],accel_mss,speed_ms,blend_radius_m)
  movel([0.518807, -1.376724, -2.573471, -0.762194, 1.570796, 2.089603],accel_mss,speed_ms,0,blend_radius_m)
  movel([0.524476, -1.392076, -2.562547, -0.757766, 1.570796, 2.095272],accel_mss,speed_ms,0,blend_radius_m)
  # End of main program
end

Machining2()
